INTERFACE ITF1

METHOD METH : BOOL
VAR_INPUT
END_VAR
END_METHOD

PROPERTY Prop : BOOL
GET
END_GET
SET
END_SET
END_PROPERTY

END_INTERFACE

(* stored: Version 1.1.0.1, ProductVersion 3.1.4024.16
   Itf ITF1: Id {e5657fdd-2b0f-433a-b7fd-718cdb622dd4}
   Method METH: Id {ac7dda20-1695-4638-a5e9-301e832555ee}
   Property Prop: Id {96b0642b-185b-4129-a7dd-5542600a5f37}
   Get Get: Id {7f04d984-ea9b-48cc-8f93-4a237996aec9}
   Set Set: Id {83ab7f49-bbbf-4304-9299-8bd6381312bb} *)
